(* Logix 5000 project; controller CIP vendor 1 type 14 code 106 rev 20.12; software revision 20.06; part 13 of 13 *)
(* tags used below, declared in another part *)
   Alarm_Present : INT[8];
   Bit : BOOL[128];
   Counter : COUNTER[10];
   IN_N7_100_199 : INT[100];
   Integer_1 : ALIAS FOR Integer[1];
   Level_Bits : BOOL[32];
   Level_Timers : TIMER[20];
   Message_Present : INT[4];
   MOA_OFF : DINT[10];
   MOA_ON : DINT[10];
   One_Shot : BOOL[128];
   OpCode_Pin : DINT[5];
   OUT_F8_0_49 : REAL[50];
   OUT_N7_0_99 : INT[100];
   Panelview : INT[40];
   PV_Message : DINT[3];
   PV_Step_Time : REAL;
   Recipe : RECIPE[41];
   SCLD_Drain_PH : REAL;
   SCLD_Dryer_Duct_Temp : REAL;
   SCLD_Dryer_Exhaust_Temp : REAL;
   SCLD_Return_Temp : REAL;
   SCLD_Rinse_Cond : REAL;
   SCLD_Solution_Tank_Lvl : REAL;
   SCLD_Supply_Flow : REAL;
   SCLD_Supply_Flow_CIP100 : REAL;
   SCLD_Supply_Flow_CIP200 : REAL;
   SCLD_Supply_Pressure : REAL;
   SCLD_Supply_Temp : REAL;
   SCLD_Wash_Chamber_Lvl : REAL;
   SCLD_Wash_Cond : REAL;
   Sequencer : CONTROL[4];
   SP_Dryer_Min_Temp : REAL;
   SP_Dryer_Temp : REAL;
   SP_Return_Temp : REAL;
   SP_Rinse_Cond : REAL;
   SP_Solution_Tank_Lvl : REAL;
   SP_Supply_Flow : REAL;
   SP_Supply_Temp : REAL;
   SP_Wash_Cond : REAL;
   SP_Wash_Cond_Hold : REAL;
   Time_Date : DINT[20];
   Timer : TIMER[99];
   Timer_Chem1_Pump : TIMER[7];
   Timer_Chem2_Pump : TIMER[7];
   Utility_Out : DINT[5];
   WashChamberDoorGasketCTRL : DINT;
(* MainProgram, continued *)

ROUTINE _89_PUMPS   (* ladder *)
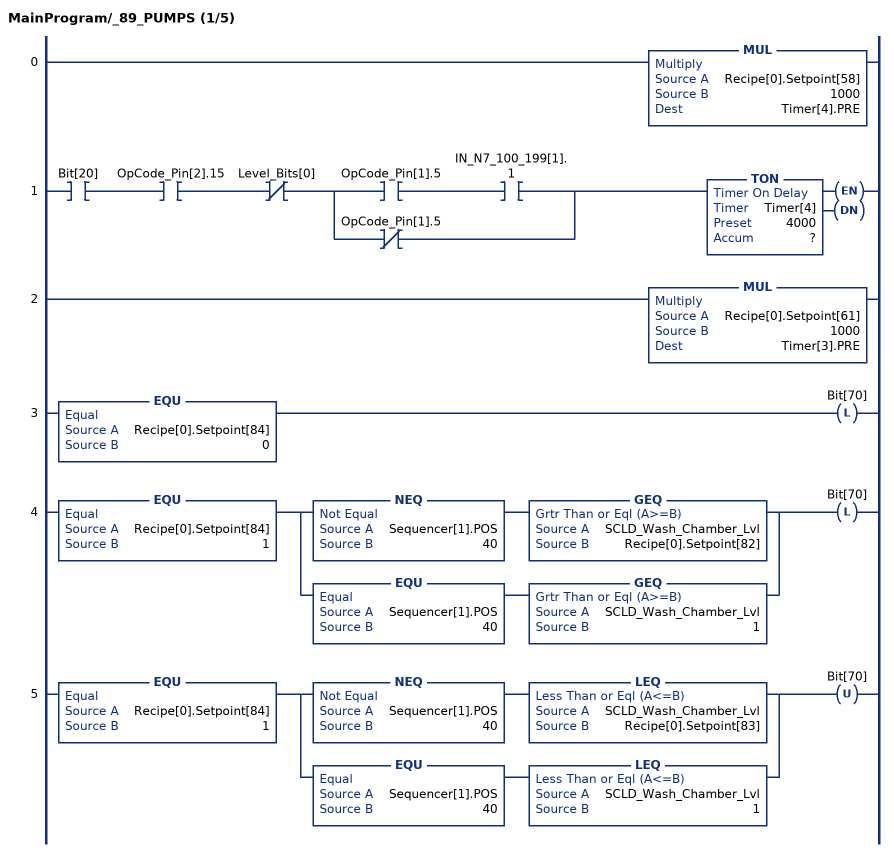
   0: MUL(Recipe[0].Setpoint[58],1000,Timer[4].PRE);
   1: XIC(Bit[20])XIC(OpCode_Pin[2].15)XIO(Level_Bits[0])[XIC(OpCode_Pin[1].5) XIC(IN_N7_100_199[1].1) ,XIO(OpCode_Pin[1].5) ]TON(Timer[4],?,?);
   2: MUL(Recipe[0].Setpoint[61],1000,Timer[3].PRE);
   3: EQU(Recipe[0].Setpoint[84],0)OTL(Bit[70]);
   4: EQU(Recipe[0].Setpoint[84],1)[NEQ(Sequencer[1].POS,40) GEQ(SCLD_Wash_Chamber_Lvl,Recipe[0].Setpoint[82]) ,EQU(Sequencer[1].POS,40) GEQ(SCLD_Wash_Chamber_Lvl,1) ]OTL(Bit[70]);
   5: EQU(Recipe[0].Setpoint[84],1)[NEQ(Sequencer[1].POS,40) LEQ(SCLD_Wash_Chamber_Lvl,Recipe[0].Setpoint[83]) ,EQU(Sequencer[1].POS,40) LEQ(SCLD_Wash_Chamber_Lvl,1) ]OTU(Bit[70]);
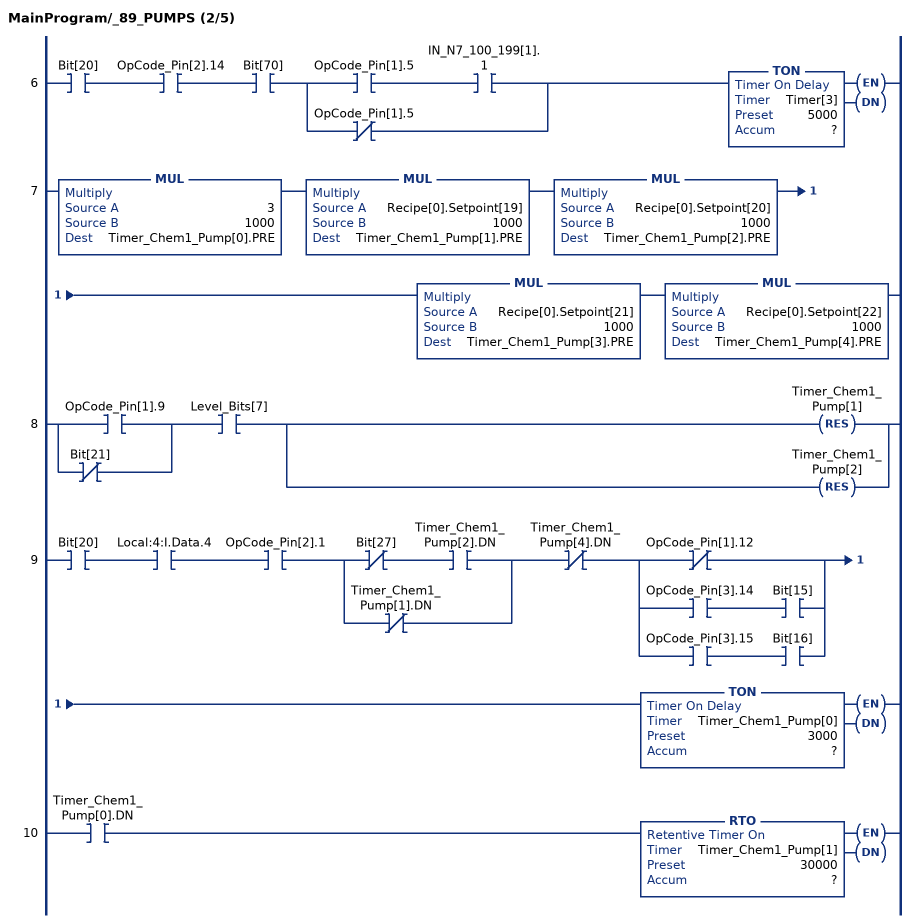
   6: XIC(Bit[20])XIC(OpCode_Pin[2].14)XIC(Bit[70])[XIC(OpCode_Pin[1].5) XIC(IN_N7_100_199[1].1) ,XIO(OpCode_Pin[1].5) ]TON(Timer[3],?,?);
   7: MUL(3,1000,Timer_Chem1_Pump[0].PRE)MUL(Recipe[0].Setpoint[19],1000,Timer_Chem1_Pump[1].PRE)MUL(Recipe[0].Setpoint[20],1000,Timer_Chem1_Pump[2].PRE)MUL(Recipe[0].Setpoint[21],1000,Timer_Chem1_Pump[3].PRE)MUL(Recipe[0].Setpoint[22],1000,Timer_Chem1_Pump[4].PRE);
   8: [XIC(OpCode_Pin[1].9) ,XIO(Bit[21]) ]XIC(Level_Bits[7])[RES(Timer_Chem1_Pump[1]) ,RES(Timer_Chem1_Pump[2]) ];
   9: XIC(Bit[20])XIC(Local:4:I.Data.4)XIC(OpCode_Pin[2].1)[XIO(Bit[27]) XIC(Timer_Chem1_Pump[2].DN) ,XIO(Timer_Chem1_Pump[1].DN) ]XIO(Timer_Chem1_Pump[4].DN)[XIO(OpCode_Pin[1].12) ,XIC(OpCode_Pin[3].14) XIC(Bit[15]) ,XIC(OpCode_Pin[3].15) XIC(Bit[16]) ]TON(Timer_Chem1_Pump[0],?,?);
   10: XIC(Timer_Chem1_Pump[0].DN)RTO(Timer_Chem1_Pump[1],?,?);
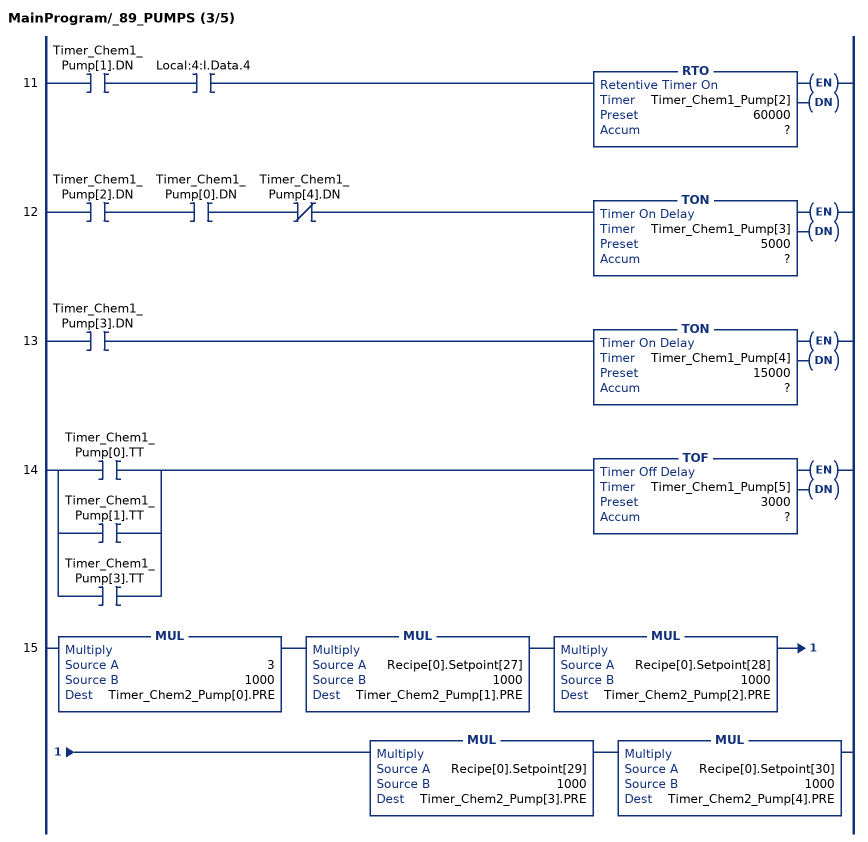
   11: XIC(Timer_Chem1_Pump[1].DN)XIC(Local:4:I.Data.4)RTO(Timer_Chem1_Pump[2],?,?);
   12: XIC(Timer_Chem1_Pump[2].DN)XIC(Timer_Chem1_Pump[0].DN)XIO(Timer_Chem1_Pump[4].DN)TON(Timer_Chem1_Pump[3],?,?);
   13: XIC(Timer_Chem1_Pump[3].DN)TON(Timer_Chem1_Pump[4],?,?);
   14: [XIC(Timer_Chem1_Pump[0].TT) ,XIC(Timer_Chem1_Pump[1].TT) ,XIC(Timer_Chem1_Pump[3].TT) ]TOF(Timer_Chem1_Pump[5],?,?);
   15: MUL(3,1000,Timer_Chem2_Pump[0].PRE)MUL(Recipe[0].Setpoint[27],1000,Timer_Chem2_Pump[1].PRE)MUL(Recipe[0].Setpoint[28],1000,Timer_Chem2_Pump[2].PRE)MUL(Recipe[0].Setpoint[29],1000,Timer_Chem2_Pump[3].PRE)MUL(Recipe[0].Setpoint[30],1000,Timer_Chem2_Pump[4].PRE);
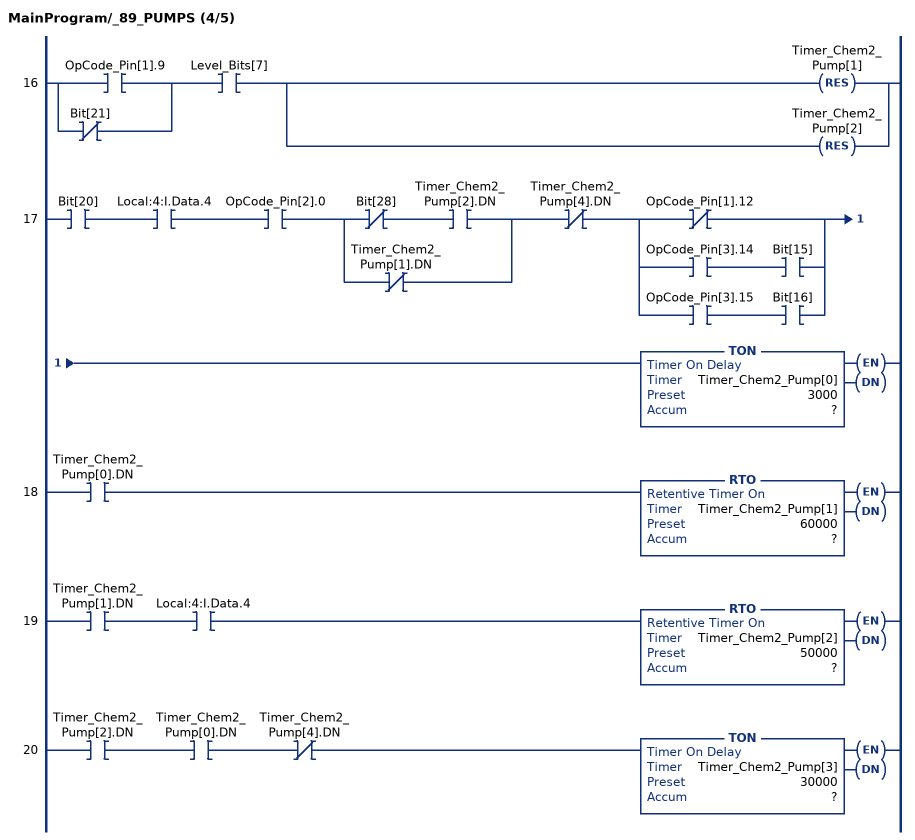
   16: [XIC(OpCode_Pin[1].9) ,XIO(Bit[21]) ]XIC(Level_Bits[7])[RES(Timer_Chem2_Pump[1]) ,RES(Timer_Chem2_Pump[2]) ];
   17: XIC(Bit[20])XIC(Local:4:I.Data.4)XIC(OpCode_Pin[2].0)[XIO(Bit[28]) XIC(Timer_Chem2_Pump[2].DN) ,XIO(Timer_Chem2_Pump[1].DN) ]XIO(Timer_Chem2_Pump[4].DN)[XIO(OpCode_Pin[1].12) ,XIC(OpCode_Pin[3].14) XIC(Bit[15]) ,XIC(OpCode_Pin[3].15) XIC(Bit[16]) ]TON(Timer_Chem2_Pump[0],?,?);
   18: XIC(Timer_Chem2_Pump[0].DN)RTO(Timer_Chem2_Pump[1],?,?);
   19: XIC(Timer_Chem2_Pump[1].DN)XIC(Local:4:I.Data.4)RTO(Timer_Chem2_Pump[2],?,?);
   20: XIC(Timer_Chem2_Pump[2].DN)XIC(Timer_Chem2_Pump[0].DN)XIO(Timer_Chem2_Pump[4].DN)TON(Timer_Chem2_Pump[3],?,?);
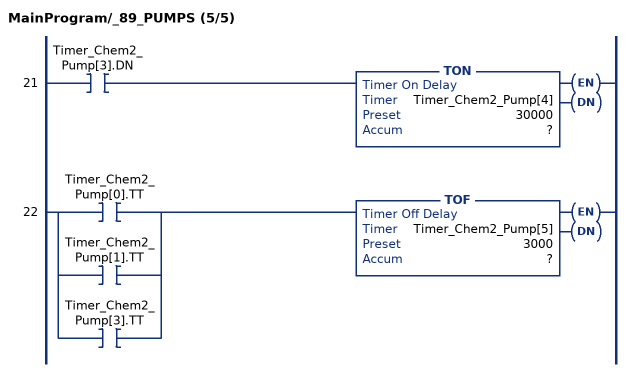
   21: XIC(Timer_Chem2_Pump[3].DN)TON(Timer_Chem2_Pump[4],?,?);
   22: [XIC(Timer_Chem2_Pump[0].TT) ,XIC(Timer_Chem2_Pump[1].TT) ,XIC(Timer_Chem2_Pump[3].TT) ]TOF(Timer_Chem2_Pump[5],?,?);
END_ROUTINE

ROUTINE _90_OUTPUTS   (* ladder *)
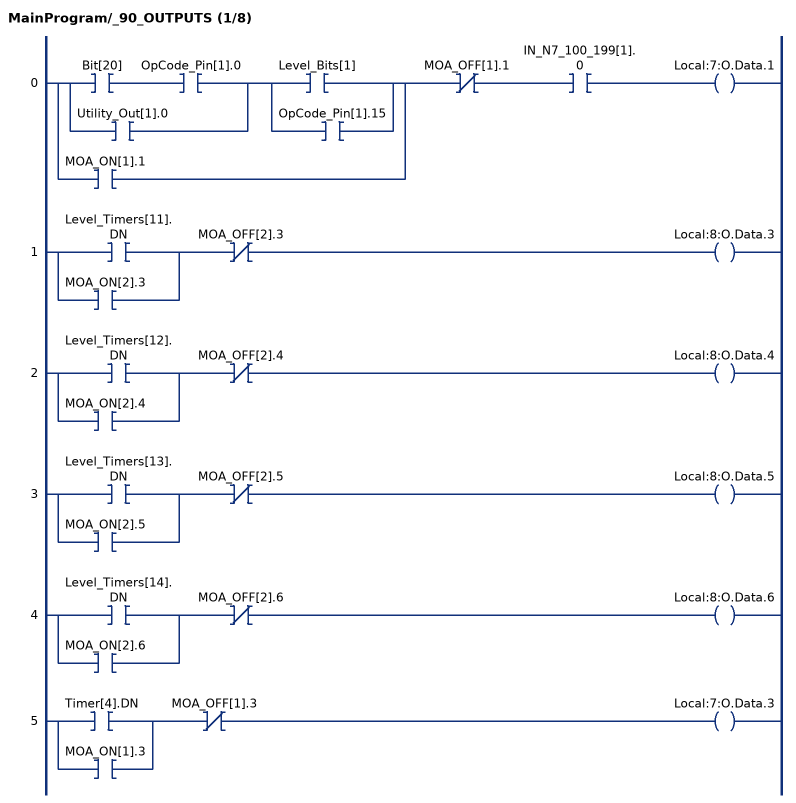
   0: [[XIC(Bit[20]) XIC(OpCode_Pin[1].0) ,XIC(Utility_Out[1].0) ] [XIC(Level_Bits[1]) ,XIC(OpCode_Pin[1].15) ] ,XIC(MOA_ON[1].1) ]XIO(MOA_OFF[1].1)XIC(IN_N7_100_199[1].0)OTE(Local:7:O.Data.1);
   1: [XIC(Level_Timers[11].DN) ,XIC(MOA_ON[2].3) ]XIO(MOA_OFF[2].3)OTE(Local:8:O.Data.3);
   2: [XIC(Level_Timers[12].DN) ,XIC(MOA_ON[2].4) ]XIO(MOA_OFF[2].4)OTE(Local:8:O.Data.4);
   3: [XIC(Level_Timers[13].DN) ,XIC(MOA_ON[2].5) ]XIO(MOA_OFF[2].5)OTE(Local:8:O.Data.5);
   4: [XIC(Level_Timers[14].DN) ,XIC(MOA_ON[2].6) ]XIO(MOA_OFF[2].6)OTE(Local:8:O.Data.6);
   5: [XIC(Timer[4].DN) ,XIC(MOA_ON[1].3) ]XIO(MOA_OFF[1].3)OTE(Local:7:O.Data.3);
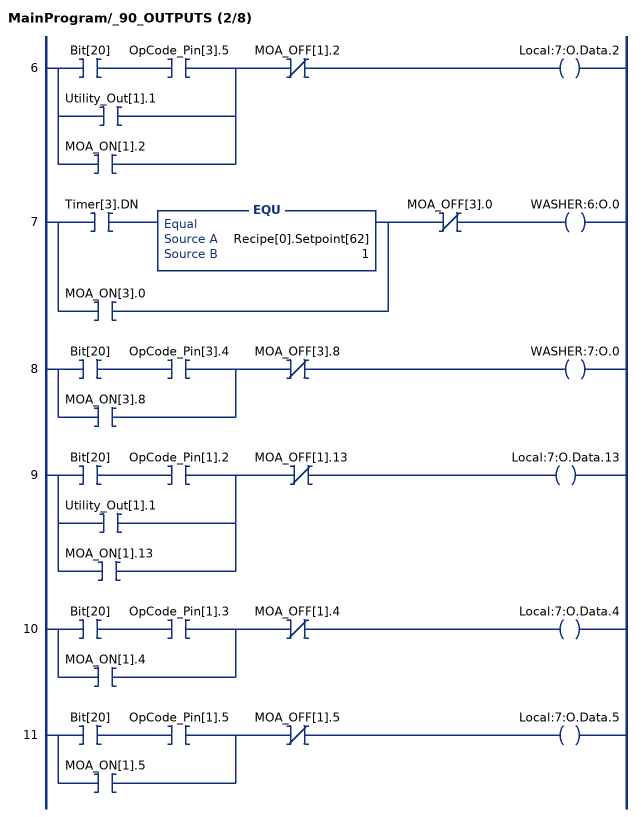
   6: [XIC(Bit[20]) XIC(OpCode_Pin[3].5) ,XIC(Utility_Out[1].1) ,XIC(MOA_ON[1].2) ]XIO(MOA_OFF[1].2)OTE(Local:7:O.Data.2);
   7: [XIC(Timer[3].DN) EQU(Recipe[0].Setpoint[62],1) ,XIC(MOA_ON[3].0) ]XIO(MOA_OFF[3].0)OTE(WASHER:6:O.0);
   8: [XIC(Bit[20]) XIC(OpCode_Pin[3].4) ,XIC(MOA_ON[3].8) ]XIO(MOA_OFF[3].8)OTE(WASHER:7:O.0);
   9: [XIC(Bit[20]) XIC(OpCode_Pin[1].2) ,XIC(Utility_Out[1].1) ,XIC(MOA_ON[1].13) ]XIO(MOA_OFF[1].13)OTE(Local:7:O.Data.13);
   10: [XIC(Bit[20]) XIC(OpCode_Pin[1].3) ,XIC(MOA_ON[1].4) ]XIO(MOA_OFF[1].4)OTE(Local:7:O.Data.4);
   11: [XIC(Bit[20]) XIC(OpCode_Pin[1].5) ,XIC(MOA_ON[1].5) ]XIO(MOA_OFF[1].5)OTE(Local:7:O.Data.5);
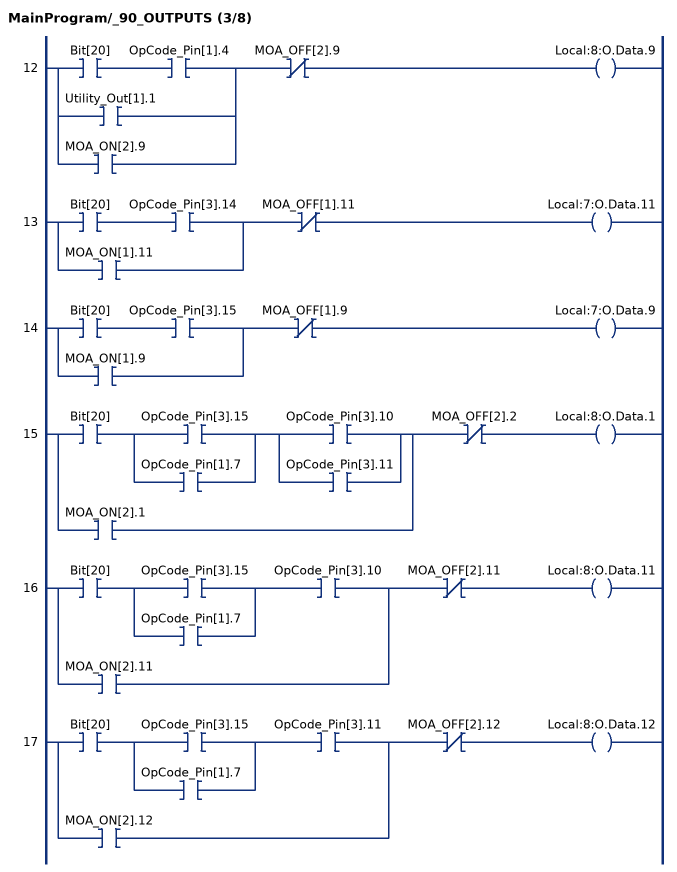
   12: [XIC(Bit[20]) XIC(OpCode_Pin[1].4) ,XIC(Utility_Out[1].1) ,XIC(MOA_ON[2].9) ]XIO(MOA_OFF[2].9)OTE(Local:8:O.Data.9);
   13: [XIC(Bit[20]) XIC(OpCode_Pin[3].14) ,XIC(MOA_ON[1].11) ]XIO(MOA_OFF[1].11)OTE(Local:7:O.Data.11);
   14: [XIC(Bit[20]) XIC(OpCode_Pin[3].15) ,XIC(MOA_ON[1].9) ]XIO(MOA_OFF[1].9)OTE(Local:7:O.Data.9);
   15: [XIC(Bit[20]) [XIC(OpCode_Pin[3].15) ,XIC(OpCode_Pin[1].7) ] [XIC(OpCode_Pin[3].10) ,XIC(OpCode_Pin[3].11) ] ,XIC(MOA_ON[2].1) ]XIO(MOA_OFF[2].2)OTE(Local:8:O.Data.1);
   16: [XIC(Bit[20]) [XIC(OpCode_Pin[3].15) ,XIC(OpCode_Pin[1].7) ] XIC(OpCode_Pin[3].10) ,XIC(MOA_ON[2].11) ]XIO(MOA_OFF[2].11)OTE(Local:8:O.Data.11);
   17: [XIC(Bit[20]) [XIC(OpCode_Pin[3].15) ,XIC(OpCode_Pin[1].7) ] XIC(OpCode_Pin[3].11) ,XIC(MOA_ON[2].12) ]XIO(MOA_OFF[2].12)OTE(Local:8:O.Data.12);
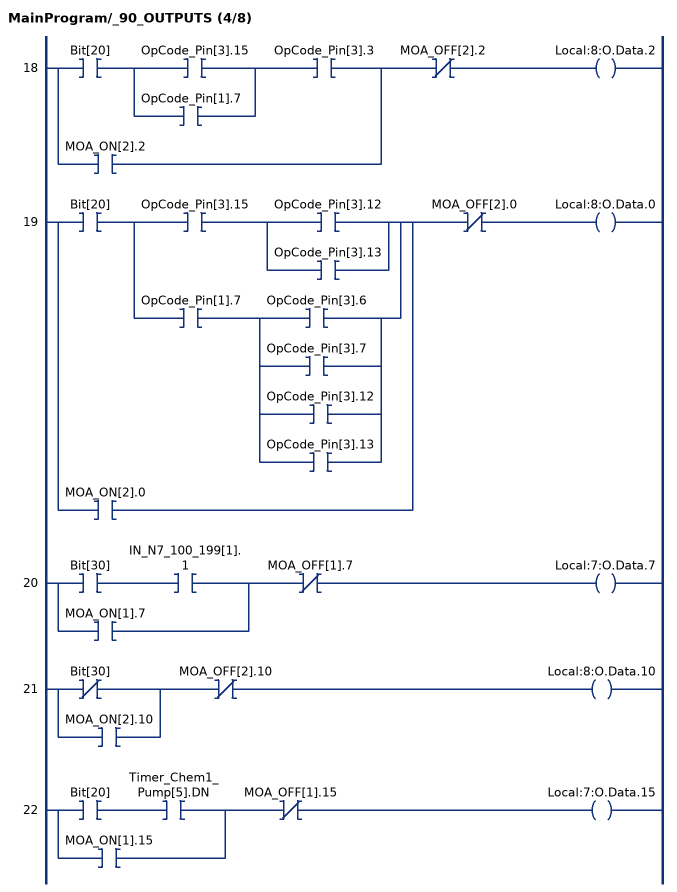
   18: [XIC(Bit[20]) [XIC(OpCode_Pin[3].15) ,XIC(OpCode_Pin[1].7) ] XIC(OpCode_Pin[3].3) ,XIC(MOA_ON[2].2) ]XIO(MOA_OFF[2].2)OTE(Local:8:O.Data.2);
   19: [XIC(Bit[20]) [XIC(OpCode_Pin[3].15) [XIC(OpCode_Pin[3].12) ,XIC(OpCode_Pin[3].13) ] ,XIC(OpCode_Pin[1].7) [XIC(OpCode_Pin[3].6) ,XIC(OpCode_Pin[3].7) ,XIC(OpCode_Pin[3].12) ,XIC(OpCode_Pin[3].13) ] ] ,XIC(MOA_ON[2].0) ]XIO(MOA_OFF[2].0)OTE(Local:8:O.Data.0);
   20: [XIC(Bit[30]) XIC(IN_N7_100_199[1].1) ,XIC(MOA_ON[1].7) ]XIO(MOA_OFF[1].7)OTE(Local:7:O.Data.7);
   21: [XIO(Bit[30]) ,XIC(MOA_ON[2].10) ]XIO(MOA_OFF[2].10)OTE(Local:8:O.Data.10);
   22: [XIC(Bit[20]) XIC(Timer_Chem1_Pump[5].DN) ,XIC(MOA_ON[1].15) ]XIO(MOA_OFF[1].15)OTE(Local:7:O.Data.15);
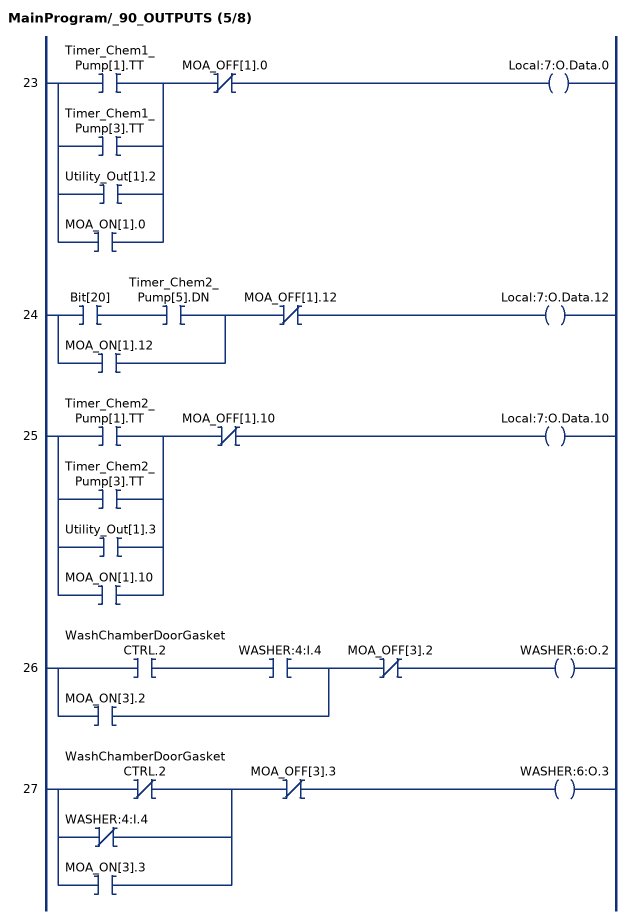
   23: [XIC(Timer_Chem1_Pump[1].TT) ,XIC(Timer_Chem1_Pump[3].TT) ,XIC(Utility_Out[1].2) ,XIC(MOA_ON[1].0) ]XIO(MOA_OFF[1].0)OTE(Local:7:O.Data.0);
   24: [XIC(Bit[20]) XIC(Timer_Chem2_Pump[5].DN) ,XIC(MOA_ON[1].12) ]XIO(MOA_OFF[1].12)OTE(Local:7:O.Data.12);
   25: [XIC(Timer_Chem2_Pump[1].TT) ,XIC(Timer_Chem2_Pump[3].TT) ,XIC(Utility_Out[1].3) ,XIC(MOA_ON[1].10) ]XIO(MOA_OFF[1].10)OTE(Local:7:O.Data.10);
   26: [XIC(WashChamberDoorGasketCTRL.2) XIC(WASHER:4:I.4) ,XIC(MOA_ON[3].2) ]XIO(MOA_OFF[3].2)OTE(WASHER:6:O.2);
   27: [XIO(WashChamberDoorGasketCTRL.2) ,XIO(WASHER:4:I.4) ,XIC(MOA_ON[3].3) ]XIO(MOA_OFF[3].3)OTE(WASHER:6:O.3);
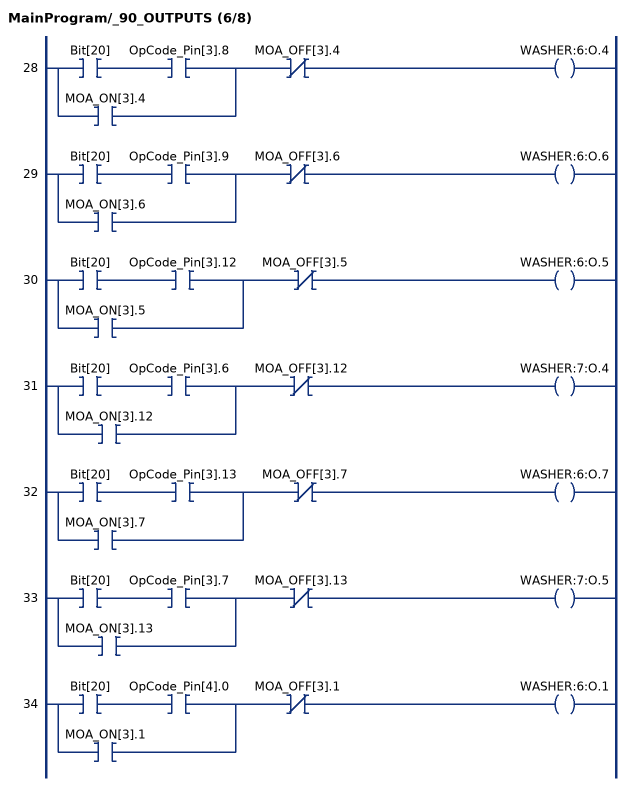
   28: [XIC(Bit[20]) XIC(OpCode_Pin[3].8) ,XIC(MOA_ON[3].4) ]XIO(MOA_OFF[3].4)OTE(WASHER:6:O.4);
   29: [XIC(Bit[20]) XIC(OpCode_Pin[3].9) ,XIC(MOA_ON[3].6) ]XIO(MOA_OFF[3].6)OTE(WASHER:6:O.6);
   30: [XIC(Bit[20]) XIC(OpCode_Pin[3].12) ,XIC(MOA_ON[3].5) ]XIO(MOA_OFF[3].5)OTE(WASHER:6:O.5);
   31: [XIC(Bit[20]) XIC(OpCode_Pin[3].6) ,XIC(MOA_ON[3].12) ]XIO(MOA_OFF[3].12)OTE(WASHER:7:O.4);
   32: [XIC(Bit[20]) XIC(OpCode_Pin[3].13) ,XIC(MOA_ON[3].7) ]XIO(MOA_OFF[3].7)OTE(WASHER:6:O.7);
   33: [XIC(Bit[20]) XIC(OpCode_Pin[3].7) ,XIC(MOA_ON[3].13) ]XIO(MOA_OFF[3].13)OTE(WASHER:7:O.5);
   34: [XIC(Bit[20]) XIC(OpCode_Pin[4].0) ,XIC(MOA_ON[3].1) ]XIO(MOA_OFF[3].1)OTE(WASHER:6:O.1);
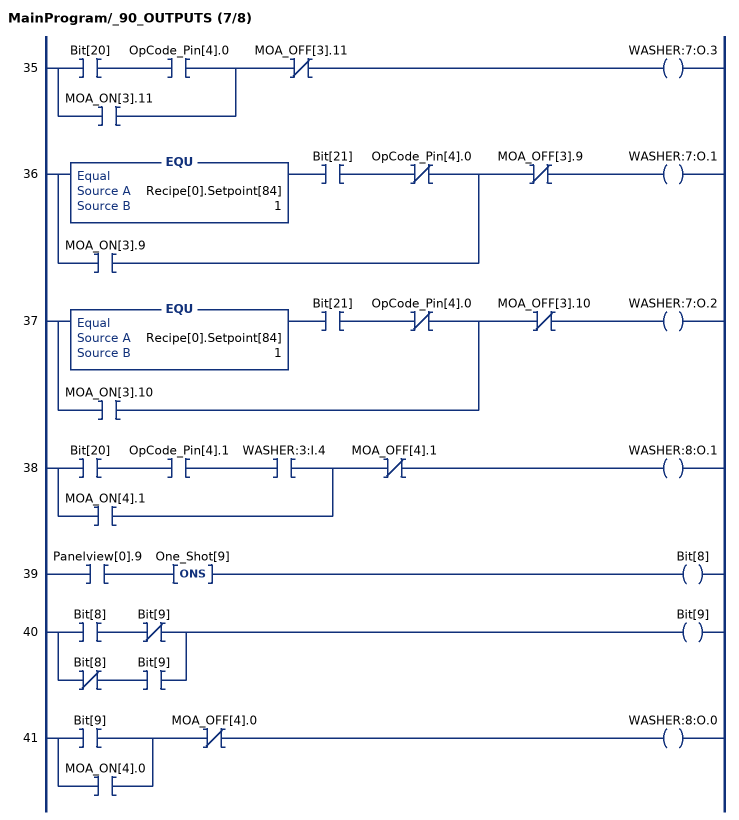
   35: [XIC(Bit[20]) XIC(OpCode_Pin[4].0) ,XIC(MOA_ON[3].11) ]XIO(MOA_OFF[3].11)OTE(WASHER:7:O.3);
   36: [EQU(Recipe[0].Setpoint[84],1) XIC(Bit[21]) XIO(OpCode_Pin[4].0) ,XIC(MOA_ON[3].9) ]XIO(MOA_OFF[3].9)OTE(WASHER:7:O.1);
   37: [EQU(Recipe[0].Setpoint[84],1) XIC(Bit[21]) XIO(OpCode_Pin[4].0) ,XIC(MOA_ON[3].10) ]XIO(MOA_OFF[3].10)OTE(WASHER:7:O.2);
   38: [XIC(Bit[20]) XIC(OpCode_Pin[4].1) XIC(WASHER:3:I.4) ,XIC(MOA_ON[4].1) ]XIO(MOA_OFF[4].1)OTE(WASHER:8:O.1);
   39: XIC(Panelview[0].9)ONS(One_Shot[9])OTE(Bit[8]);
   40: [XIC(Bit[8]) XIO(Bit[9]) ,XIO(Bit[8]) XIC(Bit[9]) ]OTE(Bit[9]);
   41: [XIC(Bit[9]) ,XIC(MOA_ON[4].0) ]XIO(MOA_OFF[4].0)OTE(WASHER:8:O.0);
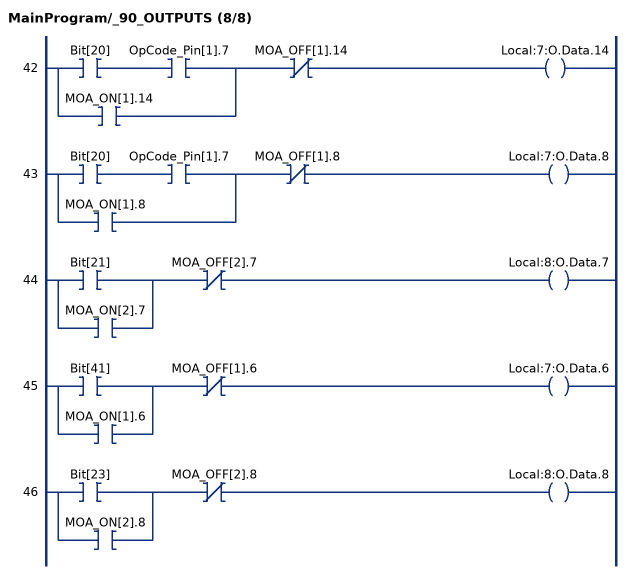
   42: [XIC(Bit[20]) XIC(OpCode_Pin[1].7) ,XIC(MOA_ON[1].14) ]XIO(MOA_OFF[1].14)OTE(Local:7:O.Data.14);
   43: [XIC(Bit[20]) XIC(OpCode_Pin[1].7) ,XIC(MOA_ON[1].8) ]XIO(MOA_OFF[1].8)OTE(Local:7:O.Data.8);
   44: [XIC(Bit[21]) ,XIC(MOA_ON[2].7) ]XIO(MOA_OFF[2].7)OTE(Local:8:O.Data.7);
   45: [XIC(Bit[41]) ,XIC(MOA_ON[1].6) ]XIO(MOA_OFF[1].6)OTE(Local:7:O.Data.6);
   46: [XIC(Bit[23]) ,XIC(MOA_ON[2].8) ]XIO(MOA_OFF[2].8)OTE(Local:8:O.Data.8);
END_ROUTINE

ROUTINE _91_SPARE_OUTPUTS   (* ladder *)
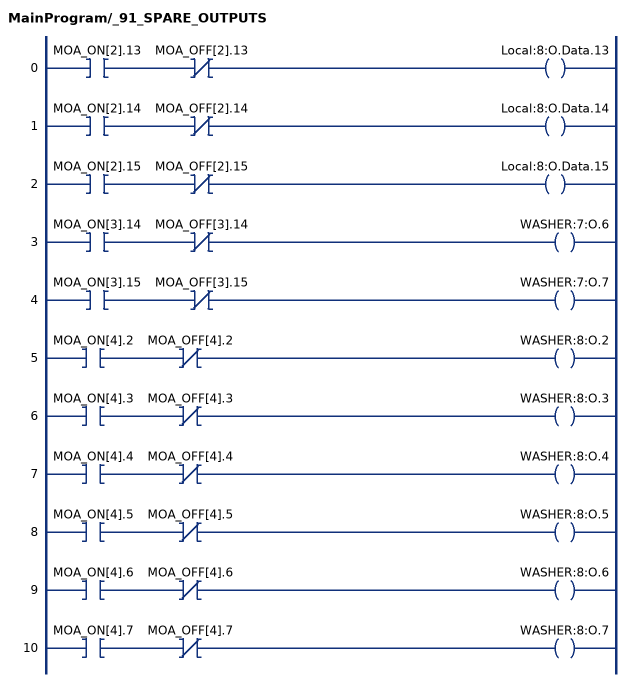
   0: XIC(MOA_ON[2].13)XIO(MOA_OFF[2].13)OTE(Local:8:O.Data.13);
   1: XIC(MOA_ON[2].14)XIO(MOA_OFF[2].14)OTE(Local:8:O.Data.14);
   2: XIC(MOA_ON[2].15)XIO(MOA_OFF[2].15)OTE(Local:8:O.Data.15);
   3: XIC(MOA_ON[3].14)XIO(MOA_OFF[3].14)OTE(WASHER:7:O.6);
   4: XIC(MOA_ON[3].15)XIO(MOA_OFF[3].15)OTE(WASHER:7:O.7);
   5: XIC(MOA_ON[4].2)XIO(MOA_OFF[4].2)OTE(WASHER:8:O.2);
   6: XIC(MOA_ON[4].3)XIO(MOA_OFF[4].3)OTE(WASHER:8:O.3);
   7: XIC(MOA_ON[4].4)XIO(MOA_OFF[4].4)OTE(WASHER:8:O.4);
   8: XIC(MOA_ON[4].5)XIO(MOA_OFF[4].5)OTE(WASHER:8:O.5);
   9: XIC(MOA_ON[4].6)XIO(MOA_OFF[4].6)OTE(WASHER:8:O.6);
   10: XIC(MOA_ON[4].7)XIO(MOA_OFF[4].7)OTE(WASHER:8:O.7);
END_ROUTINE

ROUTINE _99_DeltaV   (* ladder *)
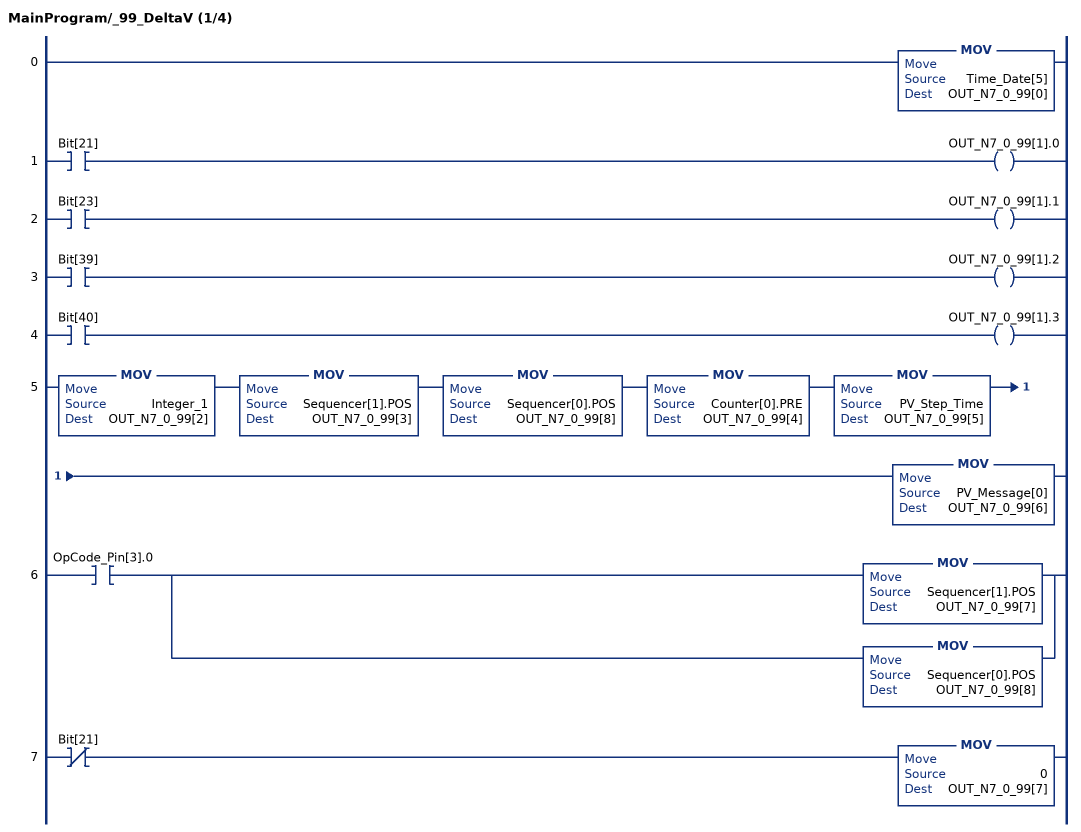
   0: MOV(Time_Date[5],OUT_N7_0_99[0]);
   1: XIC(Bit[21])OTE(OUT_N7_0_99[1].0);
   2: XIC(Bit[23])OTE(OUT_N7_0_99[1].1);
   3: XIC(Bit[39])OTE(OUT_N7_0_99[1].2);
   4: XIC(Bit[40])OTE(OUT_N7_0_99[1].3);
   5: MOV(Integer_1,OUT_N7_0_99[2])MOV(Sequencer[1].POS,OUT_N7_0_99[3])MOV(Sequencer[0].POS,OUT_N7_0_99[8])MOV(Counter[0].PRE,OUT_N7_0_99[4])MOV(PV_Step_Time,OUT_N7_0_99[5])MOV(PV_Message[0],OUT_N7_0_99[6]);
   6: XIC(OpCode_Pin[3].0)[MOV(Sequencer[1].POS,OUT_N7_0_99[7]) ,MOV(Sequencer[0].POS,OUT_N7_0_99[8]) ];
   7: XIO(Bit[21])MOV(0,OUT_N7_0_99[7]);
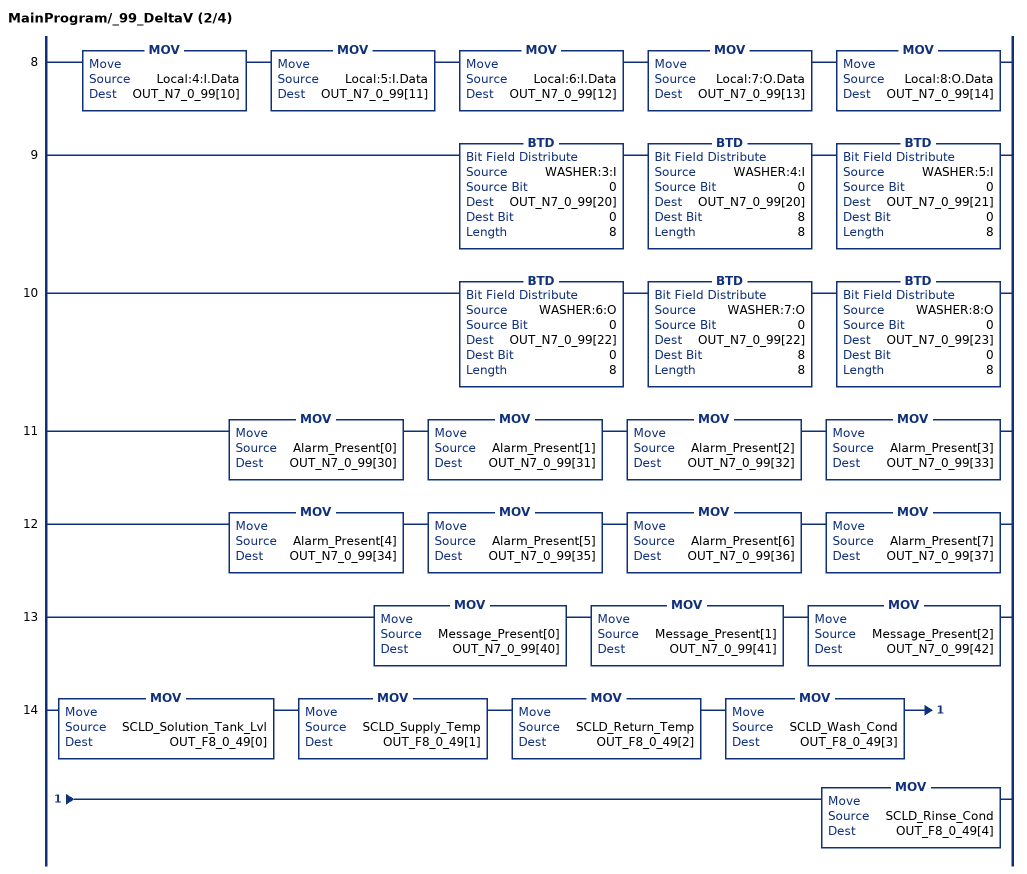
   8: MOV(Local:4:I.Data,OUT_N7_0_99[10])MOV(Local:5:I.Data,OUT_N7_0_99[11])MOV(Local:6:I.Data,OUT_N7_0_99[12])MOV(Local:7:O.Data,OUT_N7_0_99[13])MOV(Local:8:O.Data,OUT_N7_0_99[14]);
   9: BTD(WASHER:3:I,0,OUT_N7_0_99[20],0,8)BTD(WASHER:4:I,0,OUT_N7_0_99[20],8,8)BTD(WASHER:5:I,0,OUT_N7_0_99[21],0,8);
   10: BTD(WASHER:6:O,0,OUT_N7_0_99[22],0,8)BTD(WASHER:7:O,0,OUT_N7_0_99[22],8,8)BTD(WASHER:8:O,0,OUT_N7_0_99[23],0,8);
   11: MOV(Alarm_Present[0],OUT_N7_0_99[30])MOV(Alarm_Present[1],OUT_N7_0_99[31])MOV(Alarm_Present[2],OUT_N7_0_99[32])MOV(Alarm_Present[3],OUT_N7_0_99[33]);
   12: MOV(Alarm_Present[4],OUT_N7_0_99[34])MOV(Alarm_Present[5],OUT_N7_0_99[35])MOV(Alarm_Present[6],OUT_N7_0_99[36])MOV(Alarm_Present[7],OUT_N7_0_99[37]);
   13: MOV(Message_Present[0],OUT_N7_0_99[40])MOV(Message_Present[1],OUT_N7_0_99[41])MOV(Message_Present[2],OUT_N7_0_99[42]);
   14: MOV(SCLD_Solution_Tank_Lvl,OUT_F8_0_49[0])MOV(SCLD_Supply_Temp,OUT_F8_0_49[1])MOV(SCLD_Return_Temp,OUT_F8_0_49[2])MOV(SCLD_Wash_Cond,OUT_F8_0_49[3])MOV(SCLD_Rinse_Cond,OUT_F8_0_49[4]);
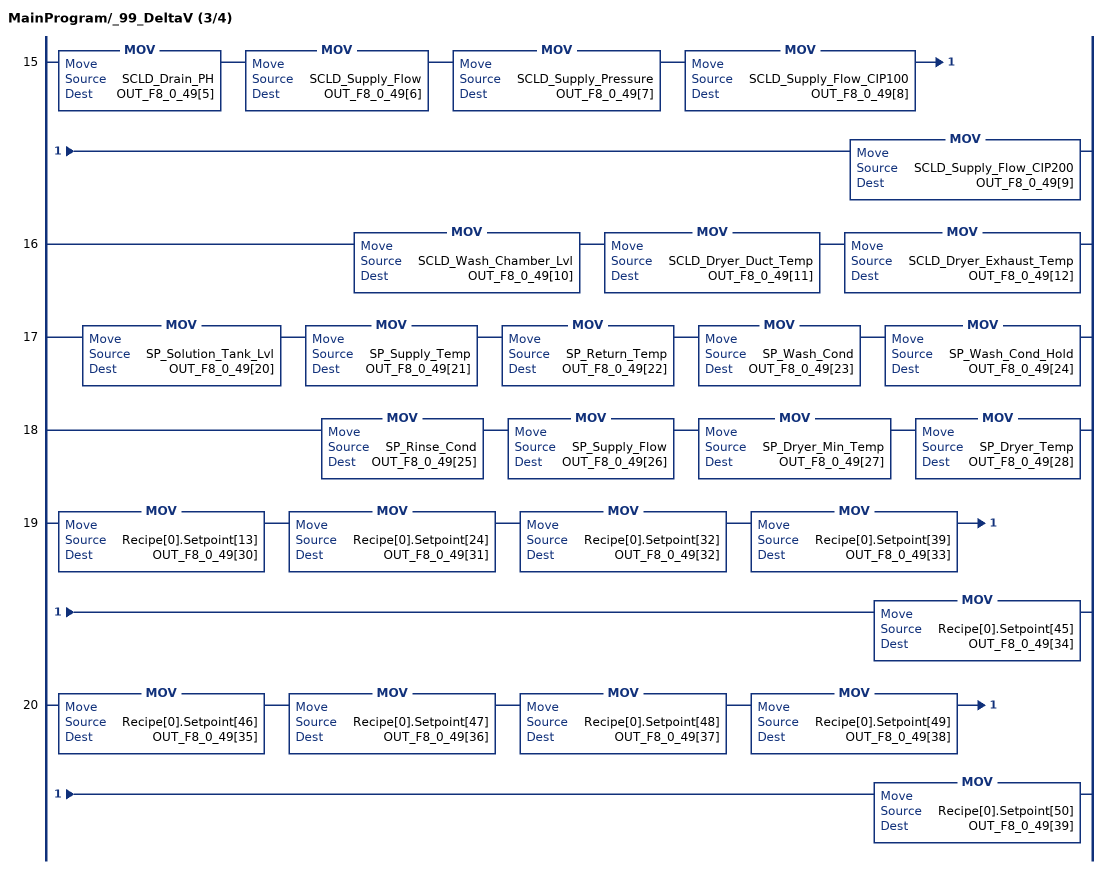
   15: MOV(SCLD_Drain_PH,OUT_F8_0_49[5])MOV(SCLD_Supply_Flow,OUT_F8_0_49[6])MOV(SCLD_Supply_Pressure,OUT_F8_0_49[7])MOV(SCLD_Supply_Flow_CIP100,OUT_F8_0_49[8])MOV(SCLD_Supply_Flow_CIP200,OUT_F8_0_49[9]);
   16: MOV(SCLD_Wash_Chamber_Lvl,OUT_F8_0_49[10])MOV(SCLD_Dryer_Duct_Temp,OUT_F8_0_49[11])MOV(SCLD_Dryer_Exhaust_Temp,OUT_F8_0_49[12]);
   17: MOV(SP_Solution_Tank_Lvl,OUT_F8_0_49[20])MOV(SP_Supply_Temp,OUT_F8_0_49[21])MOV(SP_Return_Temp,OUT_F8_0_49[22])MOV(SP_Wash_Cond,OUT_F8_0_49[23])MOV(SP_Wash_Cond_Hold,OUT_F8_0_49[24]);
   18: MOV(SP_Rinse_Cond,OUT_F8_0_49[25])MOV(SP_Supply_Flow,OUT_F8_0_49[26])MOV(SP_Dryer_Min_Temp,OUT_F8_0_49[27])MOV(SP_Dryer_Temp,OUT_F8_0_49[28]);
   19: MOV(Recipe[0].Setpoint[13],OUT_F8_0_49[30])MOV(Recipe[0].Setpoint[24],OUT_F8_0_49[31])MOV(Recipe[0].Setpoint[32],OUT_F8_0_49[32])MOV(Recipe[0].Setpoint[39],OUT_F8_0_49[33])MOV(Recipe[0].Setpoint[45],OUT_F8_0_49[34]);
   20: MOV(Recipe[0].Setpoint[46],OUT_F8_0_49[35])MOV(Recipe[0].Setpoint[47],OUT_F8_0_49[36])MOV(Recipe[0].Setpoint[48],OUT_F8_0_49[37])MOV(Recipe[0].Setpoint[49],OUT_F8_0_49[38])MOV(Recipe[0].Setpoint[50],OUT_F8_0_49[39]);
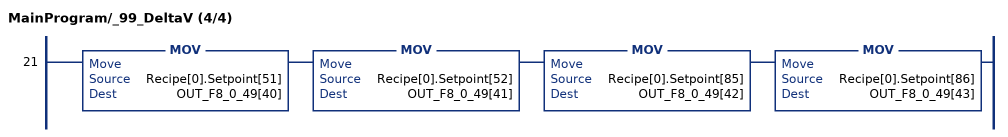
   21: MOV(Recipe[0].Setpoint[51],OUT_F8_0_49[40])MOV(Recipe[0].Setpoint[52],OUT_F8_0_49[41])MOV(Recipe[0].Setpoint[85],OUT_F8_0_49[42])MOV(Recipe[0].Setpoint[86],OUT_F8_0_49[43]);
END_ROUTINE
END_PROGRAM
